(****************************************************************************************************<br>
© Syntegon Group.<br>
All rights reserved, also regarding any disposal, exploitation, reproduction, editing, distribution,<br>
as well as in the event of applications for industrial property rights.<br>
*****************************************************************************************************<br>
DESCRIPTION:<br>
Sets or clears the fault of the whole loop: drawn red with the message while active. Faults of single<br>
movers go through m_SetMover. The fault stays until it is cleared with m_SetFault(vi_b_Active := FALSE,<br>
vi_str_Message := ''). TRUE.<br>
****************************************************************************************************)
METHOD m_SetFault : BOOL
VAR_INPUT
	vi_b_Active							: BOOL;	// TRUE: fault active
	vi_str_Message						: STRING(80);	// shown to the operator; empty shows 'Fault'
END_VAR
vo_Visu.stState.stFault.bActive := vi_b_Active;
vo_Visu.stState.stFault.sMessage := vi_str_Message;
m_SetFault := TRUE;
END_METHOD

(****************************************************************************************************<br>
© Syntegon Group.<br>
All rights reserved, also regarding any disposal, exploitation, reproduction, editing, distribution,<br>
as well as in the event of applications for industrial property rights.<br>
*****************************************************************************************************<br>
DESCRIPTION:<br>
Reports one mover at entry vi_un_Index and marks it valid. Call once per cycle per mover.<br>
*****************************************************************************************************<br>
OUTPUT VALUES:<br>
FALSE if vi_un_Index is outside the mover count set by m_SetMoverCount.<br>
****************************************************************************************************)
METHOD m_SetMover : BOOL
VAR_INPUT
	vi_un_Index							: UINT;	// [-] 0..m_SetMoverCount - 1
	vi_udn_Id							: UDINT;	// [-] unique within the loop, > 0
	vi_lr_Position						: LREAL;	// [mm] along the loop from the start of module 1 (0..m_TrackLength())
	(* Finger poses absolute in the MCS and grip states, index 0 = finger 1; entries beyond the finger count are ignored. *)
	vi_FingerStates						: ARRAY[0..VISU_GlobalConst_Param.VISU_un_MAX_FINGERS - 1] OF ST_VisuFingerState;
	vi_b_Fault							: BOOL;	// TRUE: this mover is in a fault
	vi_str_FaultMessage					: STRING(80);	// shown to the operator; empty shows 'Fault', '' without a fault
END_VAR
m_SetMover := vi_un_Index < vo_Visu.stState.nMoverCount;
IF m_SetMover THEN
	vo_Visu.stState.aMovers[vi_un_Index].nId := vi_udn_Id;
	vo_Visu.stState.aMovers[vi_un_Index].bValid := TRUE;
	vo_Visu.stState.aMovers[vi_un_Index].fPosition := vi_lr_Position;
	vo_Visu.stState.aMovers[vi_un_Index].aFingerStates := vi_FingerStates;
	vo_Visu.stState.aMovers[vi_un_Index].stFault.bActive := vi_b_Fault;
	vo_Visu.stState.aMovers[vi_un_Index].stFault.sMessage := vi_str_FaultMessage;
	vo_Visu.stState.nTimestamp := m_DcTime();
END_IF
END_METHOD

(****************************************************************************************************<br>
© Syntegon Group.<br>
All rights reserved, also regarding any disposal, exploitation, reproduction, editing, distribution,<br>
as well as in the event of applications for industrial property rights.<br>
*****************************************************************************************************<br>
DESCRIPTION:<br>
Sets how many mover entries are evaluated (limited to VISU_GlobalConst_Param.VISU_un_MAX_MOVERS); entries<br>
beyond are invalidated. TRUE if vi_un_Count fitted.<br>
****************************************************************************************************)
METHOD m_SetMoverCount : BOOL
VAR_INPUT
	vi_un_Count							: UINT;	// [-] movers
END_VAR
VAR
	un_TempIndex						: UINT;
END_VAR
m_SetMoverCount := vi_un_Count <= VISU_GlobalConst_Param.VISU_un_MAX_MOVERS;
vo_Visu.stState.nMoverCount := MIN(vi_un_Count, VISU_GlobalConst_Param.VISU_un_MAX_MOVERS);
FOR un_TempIndex := vo_Visu.stState.nMoverCount TO VISU_GlobalConst_Param.VISU_un_MAX_MOVERS - 1 DO
	vo_Visu.stState.aMovers[un_TempIndex].bValid := FALSE;
END_FOR
END_METHOD

(****************************************************************************************************<br>
© Syntegon Group.<br>
All rights reserved, also regarding any disposal, exploitation, reproduction, editing, distribution,<br>
as well as in the event of applications for industrial property rights.<br>
*****************************************************************************************************<br>
DESCRIPTION:<br>
Moves the loop's shown coordinate system (origin triad, local measuring coordinates) away from the start of<br>
the lower straight (stPose), in the loop's local frame. Geometry and mover positions stay relative to stPose.<br>
TRUE if anything changed.<br>
****************************************************************************************************)
METHOD m_SetOriginShift : BOOL
VAR_INPUT
	vi_lr_X								: LREAL;	// [mm] along the lower straight (local X)
	vi_lr_Y								: LREAL;	// [mm] along the loop's local Y, 0 = none
	vi_lr_Z								: LREAL;	// [mm] along the loop's local Z, 0 = none
END_VAR
VAR
	TempNew								: ST_VisuXtsLoopConfig;
END_VAR
TempNew := vo_Visu.stConfig;
TempNew.stOriginShift.fX := vi_lr_X;
TempNew.stOriginShift.fY := vi_lr_Y;
TempNew.stOriginShift.fZ := vi_lr_Z;
m_SetOriginShift := m_ApplyConfig(TempNew);
END_METHOD

(****************************************************************************************************<br>
© Syntegon Group.<br>
All rights reserved, also regarding any disposal, exploitation, reproduction, editing, distribution,<br>
as well as in the event of applications for industrial property rights.<br>
*****************************************************************************************************<br>
DESCRIPTION:<br>
The loop's zones for _FB_VisuZoneComponent.m_SetZone and m_ClearZones.<br>
****************************************************************************************************)
METHOD PROTECTED m_Zones : BOOL
VAR_OUTPUT
	vo_p_Count							: POINTER TO UINT;
	vo_p_Zones							: POINTER TO ARRAY[0..VISU_GlobalConst_Param.VISU_un_MAX_ZONES - 1] OF ST_VisuZone;
END_VAR
vo_p_Count := ADR(vo_Visu.stConfig.nZoneCount);
vo_p_Zones := ADR(vo_Visu.stConfig.aZones);
m_Zones := TRUE;
END_METHOD

END_FUNCTION_BLOCK

// POUs/_FC_GetVersionSynVisu
(****************************************************************************************************<br>
© Syntegon Group.<br>
All rights reserved, also regarding any disposal, exploitation, reproduction, editing, distribution,<br>
as well as in the event of applications for industrial property rights.<br>
*****************************************************************************************************<br>
DESCRIPTION:<br>
Runtime-readable version of the Syn_Visu library.<br>
*****************************************************************************************************<br>
VERSION         ¦ DATE       ¦ NAME      ¦ CHANGE<br>
Syn_Visu 3.0.0  ¦ 2026-10-31 ¦ J.Willner ¦ Naming and layout after the TCAT programming guideline<br>
Syn_Visu 3.1.0  ¦ 2026-10-31 ¦ J.Willner ¦ Faults of components and XTS movers (protocol 8)<br>
Syn_Visu 3.2.0  ¦ 2026-10-31 ¦ J.Willner ¦ _FB_VisuConveyor.m_MoveProduct<br>
Syn_Visu 3.3.0  ¦ 2026-10-31 ¦ J.Willner ¦ Zone CCS offset, origin shift per component (protocol 9)<br>
Syn_Visu 3.4.0  ¦ 2026-11-01 ¦ J.Willner ¦ m_LatchProduct: product state and robot (PLACED onto outfeeds)<br>
Syn_Visu 3.5.0  ¦ 2026-11-01 ¦ J.Willner ¦ Product shapes: box, cylinder, rounded box (protocol 10)<br>
Syn_Visu 4.0.0  ¦ 2026-11-01 ¦ J.Willner ¦ Vision system, product sensor, zones without kind (protocol 11)<br>
Syn_Visu 5.0.0  ¦ 2026-11-01 ¦ J.Willner ¦ XTS tracks of track modules, a fault per module (protocol 12)<br>
Syn_Visu 5.1.0  ¦ 2026-11-01 ¦ J.Willner ¦ Manifest sLibraryVersion: the visualisation shows the library version<br>
Syn_Visu 6.0.0  ¦ 2026-11-01 ¦ J.Willner ¦ Generic product client (nLastClientId, ePreviousState), station (protocol 13)<br>
Syn_Visu 7.0.0  ¦ 2026-11-02 ¦ J.Willner ¦ Product poses in the conveyor's coordinate system (protocol 14)<br>
Syn_Visu 7.1.0  ¦ 2026-11-05 ¦ J.Willner ¦ VISU_un_MAX_PRODUCTS 4800: registers for machines with thousands of products<br>
Syn_Visu 7.2.0  ¦ 2026-11-05 ¦ J.Willner ¦ Conveyor: product index by id, registers rearranged with MEMMOVE<br>
Syn_Visu 8.0.0  ¦ 2026-11-05 ¦ J.Willner ¦ m_Register without vi_str_Path: the symbol path comes from the instance path<br>
Syn_Visu 8.0.0  ¦ 2026-11-05 ¦ J.Willner ¦ Methods without default values: every call lists all inputs (TwinCAT 4024)<br>
Syn_Visu 9.0.0  ¦ 2026-11-05 ¦ J.Willner ¦ Zones bounded across the belt: m_SetZone vi_lr_StartY, vi_lr_EndY (protocol 15)<br>
Syn_Visu 9.1.0  ¦ 2026-11-07 ¦ J.Willner ¦ Conveyor without a body: _FB_VisuConveyor.m_SetBodyVisible (protocol 16)<br>
Syn_Visu 9.2.0  ¦ 2026-11-07 ¦ J.Willner ¦ Cartesian robot without Y or Z axis: _FB_VisuCartesian.m_SetKinematics (protocol 17)<br>
Syn_Visu 9.3.0  ¦ 2026-11-07 ¦ J.Willner ¦ Limit area for XTS gantry and Cartesian: _FB_VisuRobot.m_SetLimitArea (protocol 18)<br>
****************************************************************************************************)
FUNCTION _FC_GetVersionSynVisu : UINT
VAR_INPUT
	vi_n_VersionElement					: INT;	// [-] 1 = major, 2 = minor, 3 = revision
END_VAR

CASE vi_n_VersionElement OF
	1: _FC_GetVersionSynVisu := 9;
	2: _FC_GetVersionSynVisu := 3;
	3: _FC_GetVersionSynVisu := 0;
ELSE
	_FC_GetVersionSynVisu := 16#FFFF;
END_CASE

END_FUNCTION
